(* IEC 61131-3 sources: JingjiangMoonbox/Application/Application/任务列表/ExtTask/动作处理/动作处理 (part 3) *)

(* ---- KS_FB_SpeedControl_V2.st ---- *)
(*@CES
Name=KS_FB_SpeedControl_V2
Type=FunctionBlock
TypeGuid=6f9dac99-8de1-4efc-8465-68ac443b7d08
Guid=22870b27-c9f1-48dc-96b4-a19cd60d6746
HasDeclaration=True
HasImplementation=True
*)
{DECLARATION}
FUNCTION_BLOCK KS_FB_SpeedControl_V2
VAR_INPUT
	i_xEn: BOOL;
	i_byAutoAccDecCurve:BYTE;(*2022.4.21.231635|
							默认 按照最大直线加速度进行s处理-总时间等于直线时间+平滑时间/2
						 	1：按照直线加速时间进行s处理-不限制最大加速度@总时间=直线时间
						 	2：按照直线加速时间进行s处理-限制最大加速度@总时间=直线时间
						 	3：按照直线加速时间全程s处理-@总时间=直线时间
							4: 和默认处理方式接近|@总时间=直线时间+平滑时间|2022.12.7.1704458
							5: 自动加速使用直线加速
							6: 取消s加速段，只保留s减速段|本次加减速时间是可以保证的
							7: s加速和减速保证位移一致@总时间=平滑时间+dv/i_uiMaxVel_UseCalcAcc*界面时间;平滑时间按照界面设置(s前+s后)
							8: s加速和减速保证位移一致@总时间=平滑时间+dv/i_uiMaxVel_UseCalcAcc*界面时间;平滑时间=总时间*系数
							9: s加速和减速保证位移一致@总时间=dv/i_uiMaxVel_UseCalcAcc*界面时间;平滑时间=总时间*系数*)

	i_iMsCycle_Motion: INT;(*运动周期|*)
	i_lrTimeSec_SBegin: LREAL := 30;(*S规划前半程时间|*)
	i_lrTimeSec_SEnd: LREAL := 30;(*S规划后半程时间|*)
	i_xReCalc_Target:BOOL;
	i_piTimeSec_AccDec_AllTheWay					: POINTER TO INT; (* S加减速时间 *)
	i_rVel_Max										: REAL; (* 最大速度 *)
	i_pxFlag_ArrivedToTargetVel						: POINTER TO BOOL; (* | *)
	i_rFinalVelocity								: REAL; (* 加减速末端速度 *)
	i_prVel_Cur										: POINTER TO REAL; (* 当前速度 *)
	i_prAccDecTime_ThisTime							: POINTER TO REAL; (* 本次加减速时间 *)
	i_xFlag_PTfifofull								: BOOL; (* 允许写PT使能 *)
	i_xFlag_ManuAcc									: BOOL; (* 手动加速标志 *)
	i_xFlag_ManuDec									: BOOL; (* 手动减速标志 *)
	i_xFlag_EStoping								: BOOL; (* 急停中标志 *)
	i_xFlag_Stoping									: BOOL; (* 停机中标志 *)
	i_pxFlag_Decing									: POINTER TO BOOL; (* 减速中 *)
	i_pxFlag_Accing									: POINTER TO BOOL; (* 加速中 *)
	i_xFlag_AutoAcc									: BOOL; (* 自动减速 *)
	i_xFlag_AutoDec									: BOOL; (* 自动减速 *)
	i_xFlag_InkAccing								: BOOL; (* 空转加速中 *)
	i_iIdGSE										: INT; (* 当前运行步骤 *)
	i_xFlag_Print									: BOOL;
	i_xFlag_FastStoping								: BOOL;
	i_xFlag_Ink										: BOOL;
	(*i_apstStTravelLogRec: ARRAY [1..GC_LOG_CLASSES_MAX_NUM] OF POINTER TO StTravelLogRec; (* 2021.7.5.144816/ *)*)
(*	i_bySTime_AtLeast:BYTE;(*至少s加减速时间|默认10s*)*)(*需要删除|2023.03.02.112331*)
	i_rAux_enc_vel									: REAL;//虚拟主轴的速度//当速度到位标志触发时，直接将虚拟主轴速度给目标速度
	i_rGirth_Master: REAL;
	//2025.8.25.150143+ By Liu.yt
	i_uiMaxVel_UseCalcAcc:UINT;
	i_rSpeed_SCoeff_Type789:REAL:=0.666;
	i_xUseMaxTimeAsSBegin_InLowSpeed:BOOL;
	i_iTime_AutoAcc:INT;
	i_iTime_AutoDec:INT;
END_VAR
VAR_OUTPUT
	o_xEno: BOOL;
	o_iErNo: INT;(*0.no error\-1.bad parameters\-2.bad lrVelMax&TimeAccDec|*)
	o_diVel_Virtual_Tar: DINT;
	o_lrMax_a_S_pos: LREAL;
	o_lrTime_S : LREAL;
	o_lrJerk_SBegin: LREAL;
	o_lrJerk_SEnd: LREAL;
END_VAR
VAR

	lrVel_delta: LREAL;(*速度变化量|*)
	lrJerk_SBegin: LREAL;
	lrJerk_SEnd: LREAL;
	lrAve_a: LREAL;(*全程平均加速度|*)
	lrMax_a_S: LREAL;(*S规划的最大加速度|*)
	iNum_InflectionPts: INT;
	//lrCurr_t: LREAL;(*当前时间|*)
	//lrPrev_t: LREAL;(*前次时间|*)
	xReqTestEndVelocity: BOOL;
	lrCurCycleVelVeries: LREAL;(*当前周期速度变化量|*)
	alrInflectionPts_t: ARRAY [1..2] OF LREAL:= [2(0)];(*时间轴上的拐点位置|*)

	xFlag_MotionParamInitialized: BOOL := FALSE;(*运动参数初始化标志|*)

	rMax_a_Coeff: REAL:=1.5;
	rS_AccDecTime_Coeff:REAL;(*S加减速时间-加速占的比例*)
	rAux_enc_vel_Temp:REAL;
	rTemp_Compera_Vel: REAL := 0.000016;
	fbTRIG_ArrivedTOtar: R_TRIG;
	lrFinalVelocity : LREAL;
	rAux_enc_vel : REAL;

	//2025.8.25.112406 同步

	(*2024.6.15.103803+注释*)
	rTimeSec_SBegin: REAL;(*保证位移一致的s前时间*)
	rTimeSec_SEnd: REAL;(*保证位移一致的s后时间*)
	rDistance_AccInc: REAL;(*加速过程的位移*)
	rDistance_AccDec: REAL;(*减速过程的位移*)
	rTime_Total: REAL;(*使用的总时间*)
	rTime_SmActual: REAL;(*s的总时间*)

(*	rAllTime:REAL;
	rSTime:REAL;*)
	byCalcType: BYTE;
	(*2025.2.10.112014 单位为s@Liu.yt*)
	rTimeSec_AccDec_AllTheWay_Use:REAL;(*2024.8.30.152530*)
	lrAccDecTime_ThisTime:LREAL;(*有些指针是LREAL*)
END_VAR
{IMPLEMENTATION}
o_xEno:= i_xEn;
o_iErNo:= 0;

IF i_rGirth_Master=0 THEN
	i_rGirth_Master:= 0.5;
END_IF
IF i_rSpeed_SCoeff_Type789=0 THEN
	i_rSpeed_SCoeff_Type789:= 0.6667;
END_IF
IF i_xEn THEN
	IF i_iMsCycle_Motion>0 AND
		i_lrTimeSec_SBegin>0 AND
		i_lrTimeSec_SEnd>0 THEN
		IF i_uiMaxVel_UseCalcAcc=0 THEN
			i_uiMaxVel_UseCalcAcc:=100;
		END_IF
		//在这里处理速度到位清标志动作2023.8.17.210154

		IF NOT (i_piTimeSec_AccDec_AllTheWay^>0 AND i_rVel_Max>0) THEN
			o_iErNo:= -2;
			RETURN;
		END_IF
		fbTRIG_ArrivedTOtar(CLK:=i_pxFlag_ArrivedToTargetVel^);
		IF fbTRIG_ArrivedTOtar.Q THEN
			o_diVel_Virtual_Tar:= REAL_TO_DINT(ABS(i_rAux_enc_vel));
			o_lrMax_a_S_pos:= 1;
			o_lrTime_S:= 0;
		END_IF
		IF i_pxFlag_ArrivedToTargetVel^ OR i_xReCalc_Target THEN(*速度到位|*)
			xFlag_MotionParamInitialized:= FALSE;
			o_iErNo:= -3;
			RETURN;
		END_IF

		IF NOT xFlag_MotionParamInitialized THEN(*未初始化就在这里初始化1次|*)
			xFlag_MotionParamInitialized:= TRUE;

			(*加速时间处理@2024.7.10.144615*)
			rTimeSec_AccDec_AllTheWay_Use:=i_piTimeSec_AccDec_AllTheWay^/10.0;

			(*平均加速度(m/min/s)|*)
(*			lrAve_a:= UINT_TO_LREAL(i_uiMaxVel_UseCalcAcc)(*i_pstStGrpParam^.lrVel_Max*)/INT_TO_LREAL(i_pstStGrpParam^.iTimeSec_AccDec_AllTheWay);*)
			lrAve_a:= UINT_TO_LREAL(i_uiMaxVel_UseCalcAcc)/(rTimeSec_AccDec_AllTheWay_Use);
			(*速度变化量|*)
			lrVel_delta:= i_rFinalVelocity-i_prVel_Cur^;

			IF lrVel_delta>0 THEN(*加速*)
				IF i_prVel_Cur^<9 AND(*开始的速度小于10m/min*)
					i_rFinalVelocity<=30 THEN(*目标速度小于30m/min切换*)
					IF i_byAutoAccDecCurve=4 OR
						i_byAutoAccDecCurve=7 OR
						i_byAutoAccDecCurve=8 THEN
						i_byAutoAccDecCurve:=0;(*使用默认方式*)
					END_IF
					IF rTimeSec_AccDec_AllTheWay_Use < 30 THEN(*加速时间太短了|限制最小值*)
						rTimeSec_AccDec_AllTheWay_Use:=30;
					END_IF
				END_IF
			END_IF

			(*按照平均加速度算出该段速度变化所需要的时间\
			/*由于时间是绝对量\不能出现负值|*)
			//i_prAccDecTime_ThisTime^:= ABS(lrVel_delta/lrAve_a);
			lrAccDecTime_ThisTime:= ABS(lrVel_delta/lrAve_a);

			IF lrVel_delta<0 THEN
				lrAve_a:= -lrAve_a;

			(*2018.11.26.184729|niu.j|判断如果10米印刷停机到10米空转时，
				当前速度等于目标速度导致有加速度计算，直接输出速度到位标志
				速度变化量为0时直接退出，防止rAccDecTime_ThisTime=0,导致除0*)
			ELSIF lrVel_delta=0 THEN
				i_pxFlag_ArrivedToTargetVel^:= TRUE;
				RETURN;
			ELSE;
			END_IF

			(*s加减速时间保证前后距离一致自动获取*)
			IF i_byAutoAccDecCurve=7 OR
				i_byAutoAccDecCurve=8 OR
				i_byAutoAccDecCurve=9 THEN

				IF i_byAutoAccDecCurve=7 THEN
					byCalcType:=1;(*总时间=平滑时间+dv/i_uiMaxVel_UseCalcAcc*界面时间;平滑时间按照界面设置*)
				ELSIF i_byAutoAccDecCurve=8 THEN
					byCalcType:=2;(*总时间=平滑时间+dv/i_uiMaxVel_UseCalcAcc*界面时间;平滑时间=总时间*系数*)
				ELSIF i_byAutoAccDecCurve=9 THEN
					byCalcType:=3;(*总时间=dv/i_uiMaxVel_UseCalcAcc*界面时间;平滑时间=总时间*系数*)
				ELSE
					byCalcType:=1;
				END_IF
				(*s时间占总时间的比例*)
				IF i_rSpeed_SCoeff_Type789=0 THEN
					i_rSpeed_SCoeff_Type789:=2.0/3.0;
				END_IF
				KS_GetSTime(
					byCalcType(*byCalcType*),
					i_rSpeed_SCoeff_Type789(*i_rSpeed_SCoeff*),
					LREAL_TO_INT(i_lrTimeSec_SBegin)(*i_iTimeSa_S*),
					LREAL_TO_INT(i_lrTimeSec_SEnd)(*i_iTimeEd_S*),
					i_iTime_AutoAcc(*i_iTime_Acc*),
					i_iTime_AutoDec(*i_iTime_Dec*),
					i_uiMaxVel_UseCalcAcc(*i_iVel_GetAcceleration*),
					i_prVel_Cur^(*i_rVel_Cur*),
					i_rFinalVelocity(*i_rVel_Tar*),
					ADR(rTimeSec_SBegin)(*i_prTimeSa_S*),
					ADR(rTimeSec_SEnd)(*i_prTimeEd_S*),
					ADR(rDistance_AccInc)(*i_prDis_Sa*),
					ADR(rDistance_AccDec)(*i_prDis_Ed*),
					ADR(rTime_Total)(*i_prTime_Total*),
					ADR(rTime_SmActual)(*i_prTime_SmActual*),
					ADR(lrAccDecTime_ThisTime));(*lrAccDecTime_ThisTime此时输出的直线加速的时间@下面会重新运算*)
			ELSE(*以前的方式*)
				rTimeSec_SBegin	:=	LREAL_TO_REAL(i_lrTimeSec_SBegin);
				rTimeSec_SEnd	:=	LREAL_TO_REAL(i_lrTimeSec_SEnd);
				(*2024.05.17.181512+*)
				(*s起始和结束时间做动态切换@原则是低速使用长的s时间规划*)
				IF i_xUseMaxTimeAsSBegin_InLowSpeed THEN
					IF lrAve_a>0 THEN(*加速*)
						rTimeSec_SBegin	:=	LREAL_TO_REAL(MAX(i_lrTimeSec_SBegin,i_lrTimeSec_SEnd));
						rTimeSec_SEnd	:=	LREAL_TO_REAL(MIN(i_lrTimeSec_SBegin,i_lrTimeSec_SEnd));
					ELSE(*减速*)
						rTimeSec_SBegin	:=	LREAL_TO_REAL(MIN(i_lrTimeSec_SBegin,i_lrTimeSec_SEnd));
						rTimeSec_SEnd	:=	LREAL_TO_REAL(MAX(i_lrTimeSec_SBegin,i_lrTimeSec_SEnd));
					END_IF
				END_IF
			END_IF

			rS_AccDecTime_Coeff:=rTimeSec_SBegin/(rTimeSec_SBegin+rTimeSec_SEnd);
			IF i_byAutoAccDecCurve=1 THEN(*按照直线加速时间进行s处理-不限制最大加速度*)
				//i_pstStGrpParam^.lrAccDecTime_ThisTime:= i_pstStGrpParam^.lrAccDecTime_ThisTime;

				IF lrAccDecTime_ThisTime>(rTimeSec_SBegin+rTimeSec_SEnd) THEN(*梯形|*)
					iNum_InflectionPts:= 2;
					(*平均加速度(m/min/s)|*)
					IF lrAccDecTime_ThisTime*2<>rTimeSec_SBegin+rTimeSec_SEnd THEN
						lrMax_a_S:= 2*lrVel_delta/(2*lrAccDecTime_ThisTime-rTimeSec_SBegin-rTimeSec_SEnd);
					END_IF

					lrJerk_SBegin:= lrMax_a_S/rTimeSec_SBegin;
					lrJerk_SEnd:= lrMax_a_S/rTimeSec_SEnd;
					alrInflectionPts_t[1]:= rTimeSec_SBegin;
					alrInflectionPts_t[2]:= lrAccDecTime_ThisTime-rTimeSec_SEnd;
				ELSE(*三角形*)
					iNum_InflectionPts:= 1;
					(*平均加速度(m/min/s)|*)
					IF lrAccDecTime_ThisTime<>0 THEN
						lrMax_a_S:= 2*lrVel_delta/(lrAccDecTime_ThisTime);
					END_IF

					alrInflectionPts_t[1]:= ABS(lrAccDecTime_ThisTime*(rS_AccDecTime_Coeff));
					alrInflectionPts_t[2]:= ABS(lrAccDecTime_ThisTime*(1-rS_AccDecTime_Coeff));
(*
					lrJerk_SBegin:= lrMax_a_S/alrInflectionPts_t[1];
					lrJerk_SEnd:= lrMax_a_S/alrInflectionPts_t[2];
*)
					rTimeSec_SBegin:= LREAL_TO_REAL(alrInflectionPts_t[1]);
					rTimeSec_SEnd:= LREAL_TO_REAL(alrInflectionPts_t[2]);
					lrJerk_SBegin:= lrMax_a_S/rTimeSec_SBegin;
					lrJerk_SEnd:= lrMax_a_S/rTimeSec_SEnd;
				END_IF
			ELSIF i_byAutoAccDecCurve=2 THEN(*按照直线加速时间进行s处理-限制最大加速度|这中情况下s加减速时间会变*)
				lrAccDecTime_ThisTime:= lrAccDecTime_ThisTime;
				(*在不修改s加减速时间计算最大平均加速度(m/min/s)|*)
				IF lrAccDecTime_ThisTime>(rTimeSec_SBegin+rTimeSec_SEnd) THEN(*梯形|*)
					IF lrAccDecTime_ThisTime*2>rTimeSec_SBegin+rTimeSec_SEnd THEN
						lrMax_a_S:= 2*lrVel_delta/(2*lrAccDecTime_ThisTime-rTimeSec_SBegin-rTimeSec_SEnd);
					END_IF
				ELSE
					(*重新计算平均加速度(m/min/s)|*)
					IF lrAccDecTime_ThisTime<>0 THEN
						lrMax_a_S:= 2*lrVel_delta/(lrAccDecTime_ThisTime);
					END_IF
				END_IF

				IF ABS(lrAve_a)*rMax_a_Coeff<ABS(lrMax_a_S) THEN(*超过了我限制的最大加速度-按照最大加速度处理
													我就需要重新计算s加减速时间*)
					lrMax_a_S:=lrAve_a*rMax_a_Coeff;(*最大加速度为直线加速度的倍数*)

					(*重新计算s时间*)
					rTimeSec_SBegin:=LREAL_TO_REAL(2*(lrAccDecTime_ThisTime-ABS(lrVel_delta/lrMax_a_S))*rS_AccDecTime_Coeff);
					rTimeSec_SEnd:=LREAL_TO_REAL(2*(lrAccDecTime_ThisTime-ABS(lrVel_delta/lrMax_a_S))*(1-rS_AccDecTime_Coeff));
				END_IF

				IF lrAccDecTime_ThisTime>(rTimeSec_SBegin+rTimeSec_SEnd) THEN(*梯形|*)
					iNum_InflectionPts:= 2;

					lrJerk_SBegin:= lrMax_a_S/rTimeSec_SBegin;
					lrJerk_SEnd:= lrMax_a_S/rTimeSec_SEnd;
					alrInflectionPts_t[1]:= rTimeSec_SBegin;
					alrInflectionPts_t[2]:= lrAccDecTime_ThisTime-rTimeSec_SEnd;
				ELSE(*三角形*)
					iNum_InflectionPts:= 1;

					alrInflectionPts_t[1]:= ABS(lrAccDecTime_ThisTime*(rS_AccDecTime_Coeff));
					alrInflectionPts_t[2]:= ABS(lrAccDecTime_ThisTime*(1-rS_AccDecTime_Coeff));
(*
					lrJerk_SBegin:= lrMax_a_S/alrInflectionPts_t[1];
					lrJerk_SEnd:= lrMax_a_S/alrInflectionPts_t[2];
*)
					rTimeSec_SBegin:= LREAL_TO_REAL(alrInflectionPts_t[1]);
					rTimeSec_SEnd:= LREAL_TO_REAL(alrInflectionPts_t[2]);
					lrJerk_SBegin:= lrMax_a_S/rTimeSec_SBegin;
					lrJerk_SEnd:= lrMax_a_S/rTimeSec_SEnd;
				END_IF

			ELSIF i_byAutoAccDecCurve=3 THEN(*按照直线加速时间全程s处理*)
				(*三角形*)
				iNum_InflectionPts:= 1;
				(*平均加速度(m/min/s)|*)
				IF lrAccDecTime_ThisTime<>0 THEN
					lrMax_a_S:= 2*lrVel_delta/(lrAccDecTime_ThisTime);
				END_IF

				alrInflectionPts_t[1]:= ABS(lrAccDecTime_ThisTime*(rS_AccDecTime_Coeff));
				alrInflectionPts_t[2]:= ABS(lrAccDecTime_ThisTime*(1-rS_AccDecTime_Coeff));
(*
				lrJerk_SBegin:= lrMax_a_S/alrInflectionPts_t[1];
				lrJerk_SEnd:= lrMax_a_S/alrInflectionPts_t[2];
*)
				rTimeSec_SBegin:= LREAL_TO_REAL(alrInflectionPts_t[1]);
				rTimeSec_SEnd:= LREAL_TO_REAL(alrInflectionPts_t[2]);
				lrJerk_SBegin:= lrMax_a_S/rTimeSec_SBegin;
				lrJerk_SEnd:= lrMax_a_S/rTimeSec_SEnd;

			ELSIF i_byAutoAccDecCurve=4 OR(*强制在直线的基础时间上增加了s时间*)
					i_byAutoAccDecCurve=7 OR(*s是保证位移相等的@s按照界面设置*)
					i_byAutoAccDecCurve=8 OR(*s是保证位移相等的@s按照总时间的比例*)
					i_byAutoAccDecCurve=9 THEN(*s是保证位移相等的@保证总时间是直线计算的时间的*)

					iNum_InflectionPts:=2;(*还是使用T形方式|*)
					(*使用前后不同的S加速时间|2023.03.02.113109|*)
					lrMax_a_S:=2*lrVel_delta/(rTimeSec_SBegin+rTimeSec_SEnd+
								2*lrAccDecTime_ThisTime);

					lrAccDecTime_ThisTime:= lrAccDecTime_ThisTime+rTimeSec_SBegin+rTimeSec_SEnd;
					lrJerk_SBegin:= lrMax_a_S/rTimeSec_SBegin;
					lrJerk_SEnd:= lrMax_a_S/rTimeSec_SEnd;
					alrInflectionPts_t[1]:= rTimeSec_SBegin;
					alrInflectionPts_t[2]:= lrAccDecTime_ThisTime-rTimeSec_SEnd;

			ELSIF i_byAutoAccDecCurve=6 THEN(*取消s加速段，只保留s减速段|本次加减速时间是可以保证的*)
				//lrAccDecTime_ThisTime:= lrAccDecTime_ThisTime;

				IF lrAccDecTime_ThisTime>(rTimeSec_SEnd) THEN(*梯形|*)
					iNum_InflectionPts:= 2;
					(*平均加速度(m/min/s)|*)
					lrMax_a_S:= 2*lrVel_delta/(2*lrAccDecTime_ThisTime-rTimeSec_SEnd);

					lrJerk_SBegin:=0;
					lrJerk_SEnd:= lrMax_a_S/rTimeSec_SEnd;
					alrInflectionPts_t[1]:= 0;
					alrInflectionPts_t[2]:= lrAccDecTime_ThisTime-rTimeSec_SEnd;
				ELSE(*三角形*)
					iNum_InflectionPts:= 1;
					(*平均加速度(m/min/s)|*)
					IF lrAccDecTime_ThisTime<>0 THEN
						lrMax_a_S:= 2*lrVel_delta/(lrAccDecTime_ThisTime);
					END_IF

					alrInflectionPts_t[1]:= 0;
					alrInflectionPts_t[2]:= 0;
					rTimeSec_SBegin:=0;
					rTimeSec_SEnd:= LREAL_TO_REAL(lrAccDecTime_ThisTime);
					lrJerk_SBegin:= 0;
					lrJerk_SEnd:= lrMax_a_S/rTimeSec_SEnd;
				END_IF
			ELSE(*默认*)
				(*平均加速度(m/min/s)|*)
				IF lrAccDecTime_ThisTime*2>(rTimeSec_SBegin+rTimeSec_SEnd) THEN(*梯形|*)
					iNum_InflectionPts:= 2;
					lrAccDecTime_ThisTime:= lrAccDecTime_ThisTime+rTimeSec_SBegin/2+rTimeSec_SEnd/2;
					lrMax_a_S:= lrAve_a;
					lrJerk_SBegin:= lrMax_a_S/rTimeSec_SBegin;
					lrJerk_SEnd:= lrMax_a_S/rTimeSec_SEnd;
					alrInflectionPts_t[1]:= rTimeSec_SBegin;
					alrInflectionPts_t[2]:= lrAccDecTime_ThisTime-rTimeSec_SEnd;
				ELSE(*三角形*)
					iNum_InflectionPts:= 1;
					lrAccDecTime_ThisTime:= lrAccDecTime_ThisTime*2;
					lrMax_a_S:= lrAve_a;
					alrInflectionPts_t[1]:= lrAccDecTime_ThisTime/2;
					alrInflectionPts_t[2]:= lrAccDecTime_ThisTime/2;
					rTimeSec_SBegin:= LREAL_TO_REAL(alrInflectionPts_t[1]);
					rTimeSec_SEnd:= LREAL_TO_REAL(alrInflectionPts_t[2]);
					lrJerk_SBegin:= lrMax_a_S/rTimeSec_SBegin;
					lrJerk_SEnd:= lrMax_a_S/rTimeSec_SEnd;
				END_IF
			END_IF

			i_prAccDecTime_ThisTime^:= LREAL_TO_REAL(lrAccDecTime_ThisTime);//写入到输出

			IF i_xFlag_ManuDec OR i_xFlag_EStoping(*2023.08.28.193725*)
				OR i_xFlag_Stoping OR
				i_xFlag_FastStoping OR(*手动减速和急停/停机/快速停止中采用直线减速|*)
				(*2023.3.2.164553 空转自动减速也使用直线减速*)
				(i_xFlag_AutoDec AND (i_xflag_ink OR i_byAutoAccDecCurve=5)) THEN
					o_diVel_Virtual_Tar:= LREAL_TO_DINT(i_rFinalVelocity*GC_LRMOTORPPR/i_rGirth_Master/60.0/1000.0);
					o_lrMax_a_S_pos:= lrAve_a*GC_LRMOTORPPR/i_rGirth_Master/60.0/1000.0/1000.0;
					o_lrTime_S := 0;
					o_lrJerk_SBegin:= 0;
					o_lrJerk_SEnd:= 0;
			ELSIF i_xFlag_ManuAcc OR
				i_xFlag_InkAccing OR(*手动加速/空转加速用手动直线加速|*)
				(*2023.3.2.164553 空转自动加速使用直线加速*)
				(i_xFlag_AutoAcc AND (i_xflag_ink OR i_byAutoAccDecCurve=5)) THEN
					o_diVel_Virtual_Tar:= LREAL_TO_DINT(i_rFinalVelocity*GC_LRMOTORPPR/i_rGirth_Master/60.0/1000.0);
					o_lrMax_a_S_pos:= lrAve_a*GC_LRMOTORPPR/i_rGirth_Master/60.0/1000.0/1000.0;
					o_lrTime_S := 0;
					o_lrJerk_SBegin:= 0;
					o_lrJerk_SEnd:= 0;

			ELSIF i_xFlag_AutoAcc  OR(*自动加速或空转加速|*)
				i_xFlag_AutoDec THEN(*自动减速或默认停机|*)
					o_diVel_Virtual_Tar:= LREAL_TO_DINT(i_rFinalVelocity*GC_LRMOTORPPR/i_rGirth_Master/60.0/1000.0);
					o_lrMax_a_S_pos:= lrMax_a_S*GC_LRMOTORPPR/i_rGirth_Master/60.0/1000.0/1000.0;
					o_lrTime_S := alrInflectionPts_t[1];
					o_lrJerk_SBegin:= lrJerk_SBegin*GC_LRMOTORPPR/i_rGirth_Master/60.0/1000.0/1000.0/1000.0;
					o_lrJerk_SEnd:= lrJerk_SEnd*GC_LRMOTORPPR/i_rGirth_Master/60.0/1000.0/1000.0/1000.0;
			END_IF
		END_IF

		rAux_enc_vel_Temp:= LREAL_TO_REAL(ABS(i_rAux_enc_vel)*1000.0*60.0*i_rGirth_Master/GC_LRMOTORPPR);
		i_prVel_Cur^:= rAux_enc_vel_Temp;
		rAux_enc_vel:= ABS(i_rAux_enc_vel);
		lrFinalVelocity := LREAL_TO_DINT(i_rFinalVelocity*GC_LRMOTORPPR/i_rGirth_Master/60.0/1000.0);

		IF i_iIdGSE=GSE_ACCING OR
			i_iIdGSE=GSE_DECING THEN

			IF i_xFlag_ManuDec OR i_xFlag_EStoping
				OR i_xFlag_Stoping OR
				i_xFlag_FastStoping OR(*手动减速和急停/停机/快速停止中采用直线减速|*)
				(*2023.3.2.164553 空转自动减速也使用直线减速*)
				(i_xFlag_AutoDec AND (i_xflag_ink OR i_byAutoAccDecCurve=5)) THEN
				lrCurCycleVelVeries:= lrAve_a*(INT_TO_LREAL(i_iMsCycle_Motion)/1000);
				IF rAux_enc_vel > lrFinalVelocity + rTemp_Compera_Vel(*i_prVel_Cur^>i_rFinalVelocity+rTemp_Compera_Vel*) THEN
					i_pxFlag_Decing^:= TRUE;
					i_pxFlag_Accing^:= FALSE;
				ELSE
					i_pxFlag_Decing^:= FALSE;
					i_pxFlag_Accing^:= FALSE;
					i_prVel_Cur^:= i_rFinalVelocity;
//2023.8.17.213343到目标速度后，把目标速度再设置一次-为了防止手自动加速过程中停下并且速度同步
					o_diVel_Virtual_Tar:= LREAL_TO_DINT(i_rFinalVelocity*GC_LRMOTORPPR/i_rGirth_Master/60.0/1000.0);
					i_pxFlag_ArrivedToTargetVel^:= TRUE;
				END_IF
			(*2018.10.5.133955 | niu.j | 空转加速采用直线加速*)
			ELSIF i_xFlag_ManuAcc OR
				i_xFlag_InkAccing OR(*手动加速/空转加速用手动直线加速|*)
				(*2023.3.2.164553 空转自动加速使用直线加速*)
				(i_xFlag_AutoAcc AND (i_xflag_ink OR i_byAutoAccDecCurve=5)) THEN

				IF rAux_enc_vel < lrFinalVelocity-rTemp_Compera_Vel(*i_prVel_Cur^<i_rFinalVelocity-rTemp_Compera_Vel *)THEN
					i_pxFlag_Decing^:= FALSE;
					i_pxFlag_Accing^:= TRUE;
				ELSE
					i_pxFlag_Decing^:= FALSE;
					i_pxFlag_Accing^:= FALSE;
					i_prVel_Cur^:= i_rFinalVelocity;
					o_diVel_Virtual_Tar:= LREAL_TO_DINT(i_rFinalVelocity*GC_LRMOTORPPR/i_rGirth_Master/60.0/1000.0);
					i_pxFlag_ArrivedToTargetVel^:= TRUE;
				END_IF
			ELSIF i_xFlag_AutoAcc  OR(*自动加速或空转加速|*)
				i_xFlag_AutoDec THEN(*自动减速或默认停机|*)
				IF (((i_xFlag_AutoAcc OR i_xFlag_InkAccing) AND
						rAux_enc_vel < lrFinalVelocity-rTemp_Compera_Vel) (*i_prVel_Cur^<i_rFinalVelocity-rTemp_Compera_Vel) *)OR
					((i_xFlag_AutoDec OR i_xFlag_Stoping OR i_xFlag_FastStoping) AND
						rAux_enc_vel > lrFinalVelocity+rTemp_Compera_Vel))(*i_prVel_Cur^>i_rFinalVelocity+rTemp_Compera_Vel)) *)THEN

					IF i_xFlag_AutoAcc OR i_xFlag_InkAccing THEN
						i_pxFlag_Accing^:= TRUE;
						i_pxFlag_Decing^:= FALSE;
					ELSE
						i_pxFlag_Accing^:= FALSE;
						i_pxFlag_Decing^:= TRUE;
					END_IF
				ELSE
					i_pxFlag_Decing^:= FALSE;
					i_pxFlag_Accing^:= FALSE;
					i_pxFlag_ArrivedToTargetVel^:= TRUE;
					(*2018.8.15.095720 :| niu.j | 到目标速度后，当前速度赋值为目标速度*)
					i_prVel_Cur^:= i_rFinalVelocity;
					o_diVel_Virtual_Tar:= LREAL_TO_DINT(i_rFinalVelocity*GC_LRMOTORPPR/i_rGirth_Master/60.0/1000.0);
				END_IF
			END_IF

		END_IF

	ELSE
		o_iErNo:= -1;(*Bad parameters|*)
	END_IF
ELSE;
END_IF

(* ---- KS_FB_StdActionCtl.st ---- *)
(*@CES
Name=KS_FB_StdActionCtl
Type=FunctionBlock
TypeGuid=6f9dac99-8de1-4efc-8465-68ac443b7d08
Guid=676088f8-efac-4f69-8723-859df14a73f6
HasDeclaration=True
HasImplementation=True
*)
{DECLARATION}
FUNCTION_BLOCK KS_FB_StdActionCtl
(*2022.5.28.223230  修改流程增加快停处理
分开自动加减速和手动加减速变量
i_byActionCtlWay=0开机方式兼容预备直接到开机和预备后响铃完成按下空转进入*)
(*2023.3.2.211619 空转在速度过高状态下按下印刷 自动减速到空转速度的时间由30s修改未手动减速时间*)
(*2023.3.10.141728 空转速度过高进入印刷时候使用的时间用错了*)
(*2025.2.8.162545 急停时间按照输入时间执行,反算需要设置的急停时间实现*)
(*2025.2.10.112944 增加o_iTimeSec_AccDec_AllTheWay_0_1s输出单位修改为0.1s@解决急停快速停止*)
VAR_INPUT
	i_xEn									: BOOL;(*功能块使能*)
	i_byActionCtlWay						: BYTE;(*动作流程选择
													|0:预启动--空转--张力投入--印刷--空转--停机
													|1:预启动--空转--停机;预启动--张力投入--印刷(速度为0)--停机*)
	i_xBtnInk								: BOOL;(*空转按钮-包含了预启动响铃状态*)
	i_xBtnPrint								: BOOL;(*印刷按钮*)
	i_xBtnTension							: BOOL;(*张力投入按钮*)
	i_xBtnManuAcc							: BOOL;(*手动加速*)
	i_xBtnManuDec							: BOOL;(*手动减速*)
	i_xBtnAutoAccOrDec						: BOOL;(*自动加速减速*)
	i_xBtnStop								: BOOL;(*停止按钮*)
	i_xBtnFastStop							: BOOL;(*快速停止按钮|2022.4.9.233605*)
	i_xBtnEstop								: BOOL;(*急停按钮*)
	i_xTensionDne							: BOOL;(*张力投入完成了*)
	i_lrVel_Cur								: LREAL;(*当前速度*)
	i_lrVel_Max								: LREAL;(*允许的最大速度*)
	i_lrVel_Tar								: LREAL;(*自动目标速度*)
	i_lrVel_Ink								: LREAL;(*匀墨速度|*)
	i_iTime_Ink								: INT;(*空转时间|单位:s|*)
	i_iTime_Stop							: INT;(*停机时间|单位:s|*)
	i_iTime_FastStop						: INT;(*快速停机时间|单位:s|*)
	i_iTime_Estop							: INT;(*急停时间|单位:s|*)
(*2022.5.27.145223 加减速时间分开*)
(*
	i_iTime_AutoAccDec						: INT;(*自动加减速时间|单位:s|*)
	i_iTime_ManuAccDec						: INT;(*手动加减速时间|单位:s|*)
*)
	i_iTime_AutoAcc							: INT;(*自动加减速时间|单位:s|*)
	i_iTime_AutoDec							: INT;(*自动加减速时间|单位:s|*)
	i_iTime_ManuAcc							: INT;(*手动加减速时间|单位:s|*)
	i_iTime_ManuDec							: INT;(*手动加减速时间|单位:s|*)
	i_pxFlag_ArrivedToTargetVel				: POINTER TO BOOL;(*到达目标速度|在速度功能块中会修改该值。故在此使用指针2019.8.29.113741*)
	i_pxFlag_KeepAlarming					: POINTER TO BOOL;(*响铃|外部功能块会有操作*)
	i_xFilmAccFinish						: BOOL;(*料膜加速完成标志*)
	i_tmHold_PreStart						: TIME := T#3s; (* 开机预启动持续时间| 2022.5.27.143829*)
	i_bySpecialProcess						: BYTE;(*在基础的开机流程上增加了特殊开机方式切换标志|0:按照基础的|
																								 |1:北人的*)
	i_xBtnInk_BeiRen						: BOOL;(*空转按钮-专为北人使用|和基础流程的空转按钮定义不同|2022.5.28.234758*)
	(*2025.2.8.163015+*)
	i_xEstopTimeIsActTime					: BOOL;(*急停时间是实际时间标志@需要反算写入到速度功能块的时间*)
	i_uiMaxVel_UseCalcAcc					: UINT;(*计算加速度的最大速度值*)
	(*2025.2.13.131016+默认是这种方式*)
	i_xEstopTimeIsToMaxVel					: BOOL;(*急停时间是到达最大速度的时间标志@需要反算写入到速度功能块的时间*)
END_VAR
VAR_OUTPUT
	o_xEn									: BOOL;
	o_iIdGSE								: INT;(*状态!*)
	o_xFlag_Stop							: BOOL;(*停机标志*)
	o_xFlag_PreStart						: BOOL;(*预启动标志|从停机状态按(预)启动置位标志 色组速度达到空转速度清o_xFlag_PreStart标志,置位o_xFlag_Ink标志;当o_xFlag_Print标志有效后,*)
	o_xFlag_PreStart_Print					: BOOL;(*印刷预启动标志|用于华丰逻辑变量*)
	o_xFlag_Ink								: BOOL;(*匀墨标志|>20m/min不能联动*)
	o_xFlag_InkAccing						: BOOL;(*匀墨加速中<指0~10m/min那个加速过程>*)
	o_xFlag_Tension							: BOOL;(*张力投入标志|张力投入有效时收放料变频开始起作用|收放料就位后按印刷按钮,牵引压辊合压|o_xFlag_Print有效时张力投入不处理*)
	o_xFlag_Print							: BOOL;(*张力拉料标志有效时，按联动或印刷按钮 先压收牵(延时2s)再压放牵 印刷标志|印刷色组根据联动标志按用户指定的压辊顺序逐一延时压胶辊|胶辊压合完毕后才可置该标志有效|*)
	o_xFlag_Estop							: BOOL;(*急停标志|和停机一样要减速到0，只不过减速时间是急停时间*)
	o_xFlag_AutoAcc							: BOOL;(*自动加速*)
	o_xFlag_AutoDec							: BOOL;(*自动减速*)
	o_xFlag_ManuAcc							: BOOL;(*手动加速*)
	o_xFlag_ManuDec							: BOOL;(*手动减速*)
	o_xFlag_Accing							: BOOL;(*加速中*)
	o_xFlag_Decing							: BOOL;(*减速中*)
	o_xFlag_EStoping						: BOOL;(*正在急停中*)
	o_xFlag_Stoping							: BOOL;(*停机中*)
	o_xFlag_FastStoping						: BOOL;(*快速停机中*)
	(*o_xFlag_GotoInking						: BOOL;(*转到匀墨*)*)
	o_xTensionNotFinish						: BOOL;(*按下印刷按钮张力投入未完成输出*)
	o_xReCalc_Target						: BOOL;(*重新计算加减速动作参数,针对在切换变速过程逻辑*)
	o_xToPrintVelTooHigh					: BOOL;(*进入印刷状态时速度太高了*)
	o_rFinalVelocity						: REAL;(*目标速度*)
	o_iTimeSec_AccDec_AllTheWay				: INT;(*全程加减速所需要的秒|*)
	(*2025.2.10.110905+ 单位修改了0.1s@急停的时候需要更短*)
	o_iTimeSec_AccDec_AllTheWay_0_1s		: INT;(*输出时间单位为0.1s*)
	o_xVel_Tar_OverRange					: BOOL;(*目标速度超限值|2019.10.28.102337*)
END_VAR
VAR
	aR_TrigBtn								: ARRAY [1..10] OF R_TRIG;
	xTrigInk								: BOOL;(*空转按钮-包含了预启动响铃状态*)
	xTrigPrint								: BOOL;(*印刷按钮*)
	xTrigTension							: BOOL;(*张力投入按钮*)
	xTrigManuAcc							: BOOL;(*手动加速*)
	xTrigManuDec							: BOOL;(*手动减速*)
	xTrigAutoAccOrDec						: BOOL;(*自动加速减速*)
	xTrigStop								: BOOL;(*停止按钮*)
	xTrigFastStop							: BOOL;(*快速停止按钮|2022.4.9.233520*)
	xTrigEstop								: BOOL;(*急停按钮*)
	xInitialization							: BOOL;(*上电初始化*)
	byChangVelSts							: BYTE;(*变速时的状态	1 预启动--空转加速
																	2 手动加速
																    3 手动减速
																    4 自动加速
																    5 自动减速
																	6 印刷停机减速到空转
																	7 空转停机到0速
																	8 印刷停机减速到0速
																	9 印刷0速停机
																	10 急停减速
																	110 停止加减速
																	11 快速停止|2022.4.9.233449 增加*)
	byPreChangVelSts						: BYTE;
	xFlag_ArrivedToTarVel					: BOOL;
	xFlag_KeepAlarming						: BOOL;
	iToPrintMaxVel							: INT:=20;(*进入印刷的最大速度值*)
	lrFinalVelocity							: LREAL;(*保存目标速度值|只有在非加减速状态下才能将该值赋值给输出*)
	xFlag_InkToPrintAutoDec: BOOL;
	xAutoInkToPrint: BOOL;
	(*2022.5.28.233518 增加*)
	fbTon_PreStart							: TON;(*预启动计时器|2022.5.27.143640-*)
	xIamRdy: BOOL;

	(*2025.2.8.162509 设置的急停时间@100m/min的时间*)
	iTime_Estop_Set_0_1s: INT:=50;(*赋一个初值@单位0.1s*)
END_VAR
{IMPLEMENTATION}
(*处理按钮上升沿*)
aR_TrigBtn[1](CLK:=i_xBtnInk,Q=>xTrigInk);
aR_TrigBtn[2](CLK:=i_xBtnPrint,Q=>xTrigPrint);
aR_TrigBtn[3](CLK:=i_xBtnTension,Q=>xTrigTension);
aR_TrigBtn[4](CLK:=i_xBtnManuAcc,Q=>xTrigManuAcc);
aR_TrigBtn[5](CLK:=i_xBtnManuDec,Q=>xTrigManuDec);
aR_TrigBtn[6](CLK:=i_xBtnAutoAccOrDec,Q=>xTrigAutoAccOrDec);
aR_TrigBtn[7](CLK:=i_xBtnStop,Q=>xTrigStop);
aR_TrigBtn[8](CLK:=i_xBtnEstop,Q=>xTrigEstop);
aR_TrigBtn[9](CLK:=i_xBtnFastStop,Q=>xTrigFaststop);

IF i_xEstopTimeIsToMaxVel THEN
	(*2025.2.13.131116+ 急停时间是到达最大速度的时间标志@需要反算写入到速度功能块的时间*)
	IF xTrigEstop THEN(*有急停了@计算设置值*)
		IF i_uiMaxVel_UseCalcAcc<>0 AND i_lrVel_Max<>0 THEN
			iTime_Estop_Set_0_1s:=LREAL_TO_INT((UINT_TO_LREAL(i_uiMaxVel_UseCalcAcc)/i_lrVel_Max*i_iTime_Estop)*10);
			iTime_Estop_Set_0_1s:=ABS(iTime_Estop_Set_0_1s);
			IF iTime_Estop_Set_0_1s=0 THEN(*最小1s*)
				iTime_Estop_Set_0_1s:=10;
			END_IF
		ELSE
			iTime_Estop_Set_0_1s:=i_iTime_Estop*10;
		END_IF
	END_IF
ELSIF i_xEstopTimeIsActTime THEN
	(*2025.2.8.162401 急停的时间输入按照实际执行@这样就需要根据实际的时间反算设置时间*)
	IF xTrigEstop THEN(*有急停了@计算设置值*)
		IF i_uiMaxVel_UseCalcAcc<>0 AND i_lrVel_Cur<>0 THEN
			iTime_Estop_Set_0_1s:=LREAL_TO_INT((UINT_TO_REAL(i_uiMaxVel_UseCalcAcc)/i_lrVel_Cur*i_iTime_Estop)*10);
			iTime_Estop_Set_0_1s:=ABS(iTime_Estop_Set_0_1s);
			IF iTime_Estop_Set_0_1s=0 THEN(*最小1s*)
				iTime_Estop_Set_0_1s:=10;
			END_IF
		ELSE
			iTime_Estop_Set_0_1s:=i_iTime_Estop*10;
		END_IF
	END_IF
ELSE(*原来形式*)
	(*下面不用*)
	iTime_Estop_Set_0_1s:=i_iTime_Estop*10;
END_IF

IF i_pxFlag_KeepAlarming<>0 AND i_pxFlag_ArrivedToTargetVel<>0 THEN  ;ELSE RETURN;END_IF

xFlag_ArrivedToTarVel:=i_pxFlag_ArrivedToTargetVel^;
xFlag_KeepAlarming:=i_pxFlag_KeepAlarming^;
o_xReCalc_Target:=FALSE;
o_xEn:=i_xEn;

o_xVel_Tar_OverRange:=FALSE;
IF i_lrVel_Tar>i_lrVel_Max THEN(*2019.10.28.102110 对目标速度进行限值,并输出限速标志*)
	i_lrVel_Tar:=i_lrVel_Max;
	IF byChangVelSts=4 THEN(*自动加速时输出超限标志*)
		o_xVel_Tar_OverRange:=TRUE;
	END_IF
END_IF

(*预启动计时器|2022.5.27.145521*)
fbTon_PreStart(IN:=o_xFlag_PreStart OR o_xFlag_PreStart_Print,PT:=i_tmHold_PreStart);

IF  i_xEn THEN
	IF NOT xInitialization THEN(*上电默认停机状态*)
		xInitialization:=TRUE;
		o_xFlag_Stop:=TRUE;
	END_IF

	(*输入值是否合法|时间不能为0*)
	(*	KS_SetVarValue_NQ0(i_dwVarAdr, i_iSetValue, i_EmVarType)*)
	KS_SetVarValue_NQ0(ADR(i_iTime_Ink),100,TYPE_INT);
	KS_SetVarValue_NQ0(ADR(i_iTime_AutoAcc),100,TYPE_INT);
	KS_SetVarValue_NQ0(ADR(i_iTime_AutoDec),100,TYPE_INT);
	KS_SetVarValue_NQ0(ADR(i_iTime_ManuAcc),100,TYPE_INT);
	KS_SetVarValue_NQ0(ADR(i_iTime_ManuDec),100,TYPE_INT);
	KS_SetVarValue_NQ0(ADR(i_iTime_Stop),20,TYPE_INT);
	KS_SetVarValue_NQ0(ADR(i_iTime_Estop),2,TYPE_INT);
	(*修改为了0.1s单位@2025.2.10.113812+*)
	KS_SetVarValue_NQ0(ADR(iTime_Estop_Set_0_1s),20,TYPE_INT);
	KS_SetVarValue_NQ0(ADR(i_iTime_FastStop),20,TYPE_INT);

	(*2022.6.3.113642  在张力投入取消的时候清除标志|*)
	IF (i_xTensionDne OR NOT o_xFlag_Tension OR i_xBtnStop OR i_xBtnEstop) (*2022.11.21.151741 增加了按下停止和急停清除*)
		AND o_xTensionNotFinish THEN
		o_xTensionNotFinish:=FALSE ;
	END_IF

	IF NOT o_xFlag_Estop THEN(*非急停状态*)
		IF xTrigTension AND NOT o_xFlag_Print THEN(*张力投入|非印刷的时候才可以操作*)
			o_xFlag_Tension:=NOT o_xFlag_Tension;
		END_IF

		IF o_xFlag_Stop THEN(*停止状态*)
			o_xFlag_Estop:=i_xBtnEstop;(*急停处理*)
			IF o_xFlag_Estop THEN RETURN;END_IF(*急停直接返回*)

			IF xTrigInk THEN(*空转按钮*)
				xFlag_KeepAlarming:=TRUE;(*启动响铃信号*)
				o_xFlag_PreStart:=TRUE;(*进入预启动状态*)
			END_IF

			IF i_byActionCtlWay=1 THEN(*华丰流程*)
				IF xTrigPrint THEN(*印刷按钮*)
					IF NOT o_xFlag_PreStart THEN(*没有按下空转按钮 直接按的印刷按钮*)
						xFlag_KeepAlarming:=TRUE;(*启动响铃信号*)
						o_xFlag_PreStart_Print:=TRUE;(*进入印刷预启动状态*)
					END_IF
				END_IF
			ELSE(*都按标准流程走*)
				;
			END_IF
			o_xFlag_Stop:=NOT o_xFlag_PreStart AND NOT o_xFlag_PreStart_Print;
		ELSE(*处于非停止状态*)
			(*判断速度是否到位了,处理状态*)
			IF o_xFlag_Ink OR o_xFlag_Print THEN
				IF (xFlag_ArrivedToTarVel (*OR i_lrVel_Cur=0*))  AND byChangVelSts<>0 THEN
					CASE byChangVelSts OF
					6:(*印刷停机减速到空转*)
						o_xFlag_Print:=FALSE;
						o_xFlag_Ink:=TRUE;
					7:(*空转停机到0速*)
						o_xFlag_Stop:=TRUE;
					8:(*印刷停机减速到0速*);
					9:(*印刷0速停机*)
						o_xFlag_Stop:=TRUE;
					10:(*急停减速*)
						o_xFlag_EStop:=TRUE;
					11:(*快速停止|2022.4.9.235115*)
						o_xFlag_Stop:=TRUE;
					ELSE ;
					END_CASE
					byChangVelSts:=0;
					o_xReCalc_Target:=TRUE;(*在速度控制到位的时候使用该变量复位速度功能块的更新参数变量|防止在下面逻辑中清除
											xFlag_ArrivedToTarVel到位标志,导致参数不能更新直接进入下个变速逻辑*)

				END_IF
			END_IF

			(*2022.5.28.235413*)
			IF i_byActionCtlWay=1 THEN(*类华丰流程|还是使用原来的切换状态方式-即在响铃完成后进入下个状态*)
				xIamRdy:=NOT xFlag_KeepAlarming;(*响铃结束了|该条件有些瑕疵，但是可以用*)
			ELSE(*默认流程|*)
				IF i_bySpecialProcess=1 THEN(*北人需要在预启动响铃结束过程中按下空转*)
					IF o_xFlag_PreStart AND NOT xIamRdy THEN(*预启动|没有准备好的时候*)
						IF i_xBtnInk_BeiRen AND NOT xFlag_KeepAlarming THEN(*响铃结束了|检查北人空转按键*)
							xIamRdy:=TRUE;
						END_IF
						IF NOT xIamRdy THEN(*预备没准备好*)
							IF fbTon_PreStart.Q THEN(*预启动时间到|还么有按下|退出到停止*)
								o_xFlag_PreStart:=FALSE;
								o_xFlag_EStop:=i_xBtnEStop;
								IF NOT o_xFlag_EStop THEN o_xFlag_Stop:=TRUE; END_IF
							END_IF
						END_IF
					END_IF
				ELSE(*基础流程|预启动时间到了就可以进入下个状态了*)
					IF fbTon_PreStart.Q THEN(*预启动时间到*)
						xIamRdy:=TRUE;
					END_IF
				END_IF
			END_IF

(*			IF NOT xFlag_KeepAlarming THEN(*响铃完成了*)*)
			IF xIamRdy THEN(*可以进入下个开机状态了*)
				(*预启动状态*)
				IF o_xFlag_PreStart THEN(*预启动了，我们进入空转状态*)
					o_xFlag_PreStart:=FALSE;
					o_xFlag_Ink:=TRUE;
					xIamRdy:=FALSE;
					byChangVelSts:=1;(*进入空转加速逻辑*)
					(*2022.5.27.090554 增加*)
					o_xFlag_EStop:=i_xBtnEStop;
					IF NOT o_xFlag_EStop THEN o_xFlag_Stop:=i_xBtnStop; END_IF

					IF o_xFlag_EStop OR o_xFlag_Stop THEN
						byChangVelSts:=0;
					END_IF
				ELSIF o_xFlag_PreStart_Print THEN(*印刷预启动了*)
					IF i_xTensionDne THEN(*拉料完成*)
						o_xFlag_PreStart_Print:=FALSE;
						o_xFlag_Print:=TRUE;
						xIamRdy:=FALSE;
					ELSE
						o_xTensionNotFinish:=TRUE;
					END_IF
					(*2022.5.27.090540  移动位置*)
					o_xFlag_EStop:=i_xBtnEStop;
					IF NOT o_xFlag_EStop THEN o_xFlag_Stop:=i_xBtnStop; END_IF
				END_IF
			END_IF

			IF o_xFlag_PreStart OR o_xFlag_PreStart_Print THEN(*预启动中*)
				o_xFlag_EStop:=i_xBtnEStop;
				IF NOT o_xFlag_EStop THEN o_xFlag_Stop:=i_xBtnStop; END_IF
			END_IF

			(*启动状态*)
			IF o_xFlag_Ink THEN(*空转状态*)
				IF o_xFlag_InkAccing THEN;
				ELSE(*空转加速完成了*)
					IF i_byActionCtlWay=0 THEN(*常规流程*)
						IF (xTrigPrint OR xAutoInkToPrint) AND byChangVelSts=0 THEN(*并且按下了印刷键进入印刷状态*)
							IF i_xTensionDne THEN(*张力投入完成了 *)
								IF i_lrVel_Cur<=iToPrintMaxVel  THEN
									o_xFlag_Print:=TRUE;
									o_xFlag_Ink:=FALSE;
								ELSE(*速度太高不能进入印刷状态*)
									o_xToPrintVelTooHigh:=TRUE;
								END_IF
							ELSE
								o_xTensionNotFinish:=TRUE;
							END_IF
						END_IF
					END_IF
				END_IF
			ELSIF o_xFlag_Print THEN;
			END_IF

			(*清除进入印刷速度太高标志*)
			IF i_lrVel_Cur<=iToPrintMaxVel AND o_xToPrintVelTooHigh THEN
				o_xToPrintVelTooHigh:=FALSE;
			END_IF

			(*2019.10.9.112347增加了进入印刷状态时速度太高自动减速的逻辑|该状态可以被加速减速或者按下自动加速键取消掉*)
			IF NOT xFlag_InkToPrintAutoDec  THEN
				IF o_xToPrintVelTooHigh THEN
					IF byChangVelSts=0 THEN(*未有加减速的状态*)
						xTrigAutoAccOrDec:=TRUE;
						i_lrVel_Tar:=i_lrVel_Ink;(*减速到匀墨速度后进入印刷状态*)
						(*2023.3.10.141719*)
						(*使用自动减速时间变量i_iTime_AutoDec@之前使用成了i_iTime_AutoAcc变量*)
						i_iTime_AutoDec:=i_iTime_ManuDec(*30*);(*2023.3.2.211607 修改为了手动减速时间*)
						xFlag_InkToPrintAutoDec:=TRUE;
					END_IF
				END_IF
			ELSE
				IF NOT o_xToPrintVelTooHigh AND xFlag_ArrivedToTarVel THEN
					xFlag_InkToPrintAutoDec:=FALSE;
					xAutoInkToPrint:=TRUE;
				END_IF

				IF o_xToPrintVelTooHigh AND byChangVelSts=0 THEN(*未有加减速的状态|说明被打断了复位标志*)
					xFlag_InkToPrintAutoDec:=FALSE;
					o_xToPrintVelTooHigh:=FALSE;
				END_IF
			END_IF

			IF o_xFlag_Print THEN
				xAutoInkToPrint:=FALSE;
			END_IF

			(*加减速 停机 急停动作*)
			IF o_xFlag_Ink OR o_xFlag_Print THEN
				IF xTrigEstop THEN(*急停了*)
					IF NOT o_xFlag_EStoping THEN
						byChangVelSts:=10;
					END_IF
				ELSIF xTrigFaststop THEN(*快速停止*)
					IF NOT o_xFlag_FastStoping AND NOT  o_xFlag_EStoping THEN
						byChangVelSts:=11;(*快速停止*)
					END_IF
				ELSIF xTrigstop THEN(*停机*)
					IF NOT o_xFlag_FastStoping AND NOT o_xFlag_Stoping AND NOT  o_xFlag_EStoping THEN
						IF o_xFlag_Print THEN
							IF i_byActionCtlWay=1 THEN(*华丰流程*)
								IF i_lrVel_Cur=0 THEN
									byChangVelSts:=9;
								ELSE
									byChangVelSts:=8;
								END_IF
							ELSE
								byChangVelSts:=6;
							END_IF
						ELSE(*空转*)
							byChangVelSts:=7;
						END_IF
					END_IF
				ELSIF i_xBtnManuAcc THEN(*手动加速*)
					IF NOT o_xFlag_FastStoping AND NOT o_xFlag_Stoping AND NOT  o_xFlag_EStoping AND
(*2019.10.09.150026|niu.j|加减速多加限制料膜加速完成和空转加速完成*)
						((o_xFlag_Print AND i_xFilmAccFinish) OR (NOT o_xFlag_InkAccing AND o_xFlag_Ink)) THEN
						byChangVelSts:=2;
					END_IF
				ELSIF i_xBtnManuDec THEN(*手动减速*)
					IF NOT o_xFlag_FastStoping AND NOT o_xFlag_Stoping AND NOT  o_xFlag_EStoping AND
(*2019.10.09.150026|niu.j|加减速多加限制料膜加速完成和空转加速完成*)
						((o_xFlag_Print AND i_xFilmAccFinish) OR (NOT o_xFlag_InkAccing AND o_xFlag_Ink)) THEN

						byChangVelSts:=3;
					END_IF
				ELSIF xTrigAutoAccOrDec THEN(*自动加减速*)
					IF NOT o_xFlag_FastStoping AND NOT o_xFlag_Stoping AND NOT  o_xFlag_EStoping AND
(*2019.10.09.150026|niu.j|加减速多加限制料膜加速完成和空转加速完成*)
						((o_xFlag_Print AND i_xFilmAccFinish) OR (NOT o_xFlag_InkAccing AND o_xFlag_Ink)) THEN

						IF byChangVelSts<>4 AND byChangVelSts<>5 THEN
							IF i_lrVel_Cur<i_lrVel_Tar THEN
								byChangVelSts:=4;
							ELSIF i_lrVel_Cur>i_lrVel_Tar THEN
								byChangVelSts:=5;
							END_IF
						ELSE
							byChangVelSts:=110;(*停止自动加减速*)
						END_IF
					END_IF
				END_IF

				IF (byChangVelSts=2 AND NOT i_xBtnManuAcc) OR
					(byChangVelSts=3 AND NOT i_xBtnManuDec) THEN
					byChangVelSts:=110;
				END_IF

				(*复位标志*)
				o_xFlag_InkAccing:=FALSE;
			(*	o_xFlag_GotoInking:=FALSE;*)
				o_xFlag_EStoping:=FALSE;
				o_xFlag_Stoping:=FALSE;
				o_xFlag_FastStoping:=FALSE;(*2022.4.9.233906*)
				o_xFlag_AutoAcc:=FALSE;
				o_xFlag_AutoDec:=FALSE;
				o_xFlag_ManuAcc:=FALSE;
				o_xFlag_ManuDec:=FALSE;

				CASE byChangVelSts OF
					1:(*预启动--空转加速*);
						xFlag_ArrivedToTarVel:=FALSE;(*进入空转加减速逻辑*)
						o_xFlag_InkAccing:=TRUE;
						o_iTimeSec_AccDec_AllTheWay:=i_iTime_Ink;
						lrFinalVelocity:=i_lrVel_Ink;
					2:(*手动加速*)
						IF NOT xFlag_ArrivedToTarVel THEN
							IF byChangVelSts<>byPreChangVelSts AND byPreChangVelSts<>0 THEN(*状态发生了切换*)
								o_xReCalc_Target:=TRUE;
							END_IF
						ELSE
							xFlag_ArrivedToTarVel:=FALSE;(*进入手动加速逻辑*)
						END_IF
						o_xFlag_ManuAcc:=TRUE;
						o_iTimeSec_AccDec_AllTheWay:=i_iTime_ManuAcc;
						lrFinalVelocity:=i_lrVel_Max;
					3:(*手动减速*)
						IF NOT xFlag_ArrivedToTarVel THEN
							IF byChangVelSts<>byPreChangVelSts AND byPreChangVelSts<>0 THEN(*状态发生了切换*)
								o_xReCalc_Target:=TRUE;
							END_IF
						ELSE
							xFlag_ArrivedToTarVel:=FALSE;(*进入手动减速逻辑*)
						END_IF

						o_xFlag_ManuDec:=TRUE;
						o_iTimeSec_AccDec_AllTheWay:=i_iTime_ManuDec;
						lrFinalVelocity:=0;
					4:(*自动加速*)
						IF NOT xFlag_ArrivedToTarVel THEN
							IF byChangVelSts<>byPreChangVelSts AND byPreChangVelSts<>0 THEN(*状态发生了切换*)
								o_xReCalc_Target:=TRUE;
							END_IF
						ELSE
							xFlag_ArrivedToTarVel:=FALSE;(*进入自动加速逻辑*)
						END_IF
						o_xFlag_AutoAcc:=TRUE;
						o_iTimeSec_AccDec_AllTheWay:=i_iTime_AutoAcc;
						lrFinalVelocity:=i_lrVel_Tar;
					5:(*自动减速*)
						IF NOT xFlag_ArrivedToTarVel THEN
							IF byChangVelSts<>byPreChangVelSts AND byPreChangVelSts<>0 THEN(*状态发生了切换*)
								o_xReCalc_Target:=TRUE;
							END_IF
						ELSE
							xFlag_ArrivedToTarVel:=FALSE;(*进入自动减速逻辑*)
						END_IF
						o_xFlag_AutoDec:=TRUE;
						o_iTimeSec_AccDec_AllTheWay:=i_iTime_AutoDec;
						lrFinalVelocity:=i_lrVel_Tar;
					6:(*印刷停机减速到空转*)
						IF NOT xFlag_ArrivedToTarVel THEN
							IF byChangVelSts<>byPreChangVelSts AND byPreChangVelSts<>0 THEN(*状态发生了切换*)
								o_xReCalc_Target:=TRUE;
							END_IF
						ELSE
							xFlag_ArrivedToTarVel:=FALSE;(*进入停止减速逻辑*)
						END_IF
						(*o_xFlag_GotoInking:=TRUE;*)

(*						o_xFlag_AutoDec:=TRUE;*)
						o_xFlag_Stoping:=TRUE;(*2022.4.10.002820 修改为停止中*)
						o_iTimeSec_AccDec_AllTheWay:=i_iTime_Stop;
						(*2022.1.26.101627 在当前速度小于空转速度的时候保持当前速度*)
						lrFinalVelocity:=i_lrVel_Ink;
						IF i_lrVel_Cur<=i_lrVel_Ink THEN
							lrFinalVelocity:=i_lrVel_Cur;
						END_IF
					7:(*空转停机到0速*)
						IF NOT xFlag_ArrivedToTarVel THEN
							IF byChangVelSts<>byPreChangVelSts AND byPreChangVelSts<>0 THEN(*状态发生了切换*)
								o_xReCalc_Target:=TRUE;
							END_IF
						ELSE
							xFlag_ArrivedToTarVel:=FALSE;(*进入停止减速逻辑*)
						END_IF
						o_xFlag_Stoping:=TRUE;
						o_iTimeSec_AccDec_AllTheWay:=i_iTime_Stop;
						lrFinalVelocity:=0;
						IF i_lrVel_Cur=0 THEN
							xFlag_ArrivedToTarVel:=TRUE;
						END_IF
					8:(*印刷停机减速到0速*)
						IF NOT xFlag_ArrivedToTarVel THEN
							IF byChangVelSts<>byPreChangVelSts AND byPreChangVelSts<>0 THEN(*状态发生了切换*)
								o_xReCalc_Target:=TRUE;
							END_IF
						ELSE
							xFlag_ArrivedToTarVel:=FALSE;(*进入停止减速逻辑*)
						END_IF
						o_xFlag_Stoping:=TRUE;
						o_iTimeSec_AccDec_AllTheWay:=i_iTime_Stop;
						lrFinalVelocity:=0;
					9:;(*印刷0速停机*)
						IF i_lrVel_Cur=0 THEN
							xFlag_ArrivedToTarVel:=TRUE;
						END_IF
					10:(*急停减速*)
						IF NOT xFlag_ArrivedToTarVel THEN
							IF byChangVelSts<>byPreChangVelSts AND byPreChangVelSts<>0 THEN(*状态发生了切换*)
								o_xReCalc_Target:=TRUE;
							END_IF
						ELSE
							xFlag_ArrivedToTarVel:=FALSE;(*进入急停减速逻辑*)
						END_IF
						o_xFlag_EStoping:=TRUE;
						o_iTimeSec_AccDec_AllTheWay:=i_iTime_Estop;
						lrFinalVelocity:=0;
						IF i_lrVel_Cur=0 THEN
							xFlag_ArrivedToTarVel:=TRUE;
						END_IF
					11:(*2022.4.9.234241  快速停止|*)
						IF NOT xFlag_ArrivedToTarVel THEN
							IF byChangVelSts<>byPreChangVelSts AND byPreChangVelSts<>0 THEN(*状态发生了切换*)
								o_xReCalc_Target:=TRUE;
							END_IF
						ELSE
							xFlag_ArrivedToTarVel:=FALSE;(*进入停止减速逻辑*)
						END_IF
						o_xFlag_FastStoping:=TRUE;
						o_iTimeSec_AccDec_AllTheWay:=i_iTime_FastStop;
						lrFinalVelocity:=0;

						IF i_lrVel_Cur=0 THEN
							xFlag_ArrivedToTarVel:=TRUE;
						END_IF
					110:(*停止加减速*)
						xFlag_ArrivedToTarVel:=TRUE;(*停止加减速*)
				ELSE byChangVelSts:=0;
				END_CASE
			END_IF
			byPreChangVelSts:=byChangVelSts;
		END_IF
	ELSE(*急停了*)
		o_xFlag_Estop:=i_xBtnEstop;(*没有急停信号时退出该分支*)
		o_xFlag_Stop:=NOT o_xFlag_Estop;
		o_xFlag_Tension:=FALSE;
	END_IF

	IF (NOT o_xFlag_Accing AND NOT o_xFlag_Decing) OR o_xReCalc_Target THEN(*非加减速或者更新速度参数时更新目标速度*)
		o_rFinalVelocity:=LREAL_TO_REAL(lrFinalVelocity);
	END_IF

	o_xFlag_Accing:=o_xFlag_ManuAcc OR o_xFlag_AutoAcc OR o_xFlag_InkAccing;
	o_xFlag_Decing:=o_xFlag_EStoping OR o_xFlag_Stoping OR o_xFlag_FastStoping OR o_xFlag_ManuDec OR o_xFlag_AutoDec;
END_IF

(*对加减速时间进行非零保护*)
IF o_iTimeSec_AccDec_AllTheWay=0 THEN(*100S*)
	o_iTimeSec_AccDec_AllTheWay:=100;
END_IF
IF o_iTimeSec_AccDec_AllTheWay_0_1s=0 THEN(*100S*)
	o_iTimeSec_AccDec_AllTheWay_0_1s:=1000;
END_IF
(*2025.2.10.111017 该值的输出修改为了ms@为了解决急停快速停止的问题*)
IF i_xEstopTimeIsActTime OR
	i_xEstopTimeIsToMaxVel THEN
	IF o_xFlag_EStoping THEN
		o_iTimeSec_AccDec_AllTheWay_0_1s:=iTime_Estop_Set_0_1s;
	ELSE
		o_iTimeSec_AccDec_AllTheWay_0_1s:=o_iTimeSec_AccDec_AllTheWay*10;
	END_IF
ELSE(*原方式的时候统一*10*)
	o_iTimeSec_AccDec_AllTheWay_0_1s:=o_iTimeSec_AccDec_AllTheWay*10;
END_IF

(*急停停机状态以及功能块未使能时候 清除若干变量*)
IF o_xFlag_Estop OR o_xFlag_Stop OR NOT i_xEn THEN
	xFlag_ArrivedToTarVel:=TRUE;(*默认将该值写成有效 在速度功能块中不会进入加减速逻辑*)
	xFlag_KeepAlarming:=FALSE;
	xFlag_InkToPrintAutoDec:=FALSE;
	xAutoInkToPrint:=FALSE;
	o_xFlag_PreStart:=FALSE;
	o_xFlag_PreStart_Print:=FALSE;
	o_xFlag_Ink:=FALSE;
	o_xFlag_InkAccing:=FALSE;
	o_xFlag_Print:=FALSE;
	o_xFlag_AutoAcc:=FALSE;
	o_xFlag_AutoDec:=FALSE;
	o_xFlag_ManuAcc:=FALSE;
	o_xFlag_ManuDec:=FALSE;
	o_xFlag_Accing:=FALSE;
	o_xFlag_Decing:=FALSE;
	o_xFlag_Stoping:=FALSE;
	o_xFlag_FastStoping:=FALSE;
	o_xFlag_EStoping:=FALSE;
	(*o_xFlag_GotoInking:=FALSE;*)
	o_xTensionNotFinish:=FALSE;
	o_xToPrintVelTooHigh:=FALSE;
	lrFinalVelocity:=0;
	o_rFinalVelocity:=0;
	byChangVelSts:=0;
	byPreChangVelSts:=0;
	xIamRdy:=FALSE;(*2022.5.28.234611*)
	fbTon_PreStart(IN:=FALSE);
	IF NOT i_xEn THEN
		o_iIdGSE:=GSE_UNKNOWN;
		o_xFlag_Estop:=FALSE;
		o_xFlag_Stop:=FALSE;
		o_xFlag_Tension:=FALSE;
	END_IF
END_IF

i_pxFlag_ArrivedToTargetVel^:=xFlag_ArrivedToTarVel;
i_pxFlag_KeepAlarming^:=xFlag_KeepAlarming;

(*输出以前逻辑所需要的状态*)
o_iIdGSE:=GSE_UNKNOWN;
IF o_xFlag_Estop THEN
	o_iIdGSE:=GSE_ESTOP;
ELSIF o_xFlag_Stop THEN
	o_iIdGSE:=GSE_STOP;
ELSIF o_xFlag_Accing THEN
	o_iIdGSE:=GSE_ACCING;
ELSIF o_xFlag_Decing THEN
	o_iIdGSE:=GSE_DECING;
ELSIF o_xFlag_Ink THEN
	o_iIdGSE:=GSE_INK;
ELSIF o_xFlag_Print THEN
	o_iIdGSE:=GSE_PRINT;
ELSIF o_xFlag_PreStart THEN
	o_iIdGSE:=GSE_PRESTART;
ELSIF o_xFlag_PreStart_Print THEN
	o_iIdGSE:=GSE_PRINT_PRESTART;
ELSIF o_xFlag_Tension THEN
	o_iIdGSE:=GSE_KEEP_TENSION;
END_IF
